(* Logix 5000 project; controller R400_500_XLS vendor 1 type 14 code 216 rev 31.11; software revision 31.01; part 9 of 32 *)
(* tags used below, declared in another part *)
   Abort1 : DINT;   // Not Used
   Alarm : SINT;   // Wait 3 seconds
   Ashutdown : SINT;   // Not Used
   Condenser : INT;
   CondenserHighFlow_1 : BOOL;   // Enables the condenser high flow valve
   CondenserHighFlow_2 : BOOL;   // Enables the condenser high flow valve
   CondenserLowFlow_1 : BOOL;   // Enables the condenser low flow valve
   CondenserLowFlow_2 : BOOL;   // Enables the condenser low flow valve
   CURRENT_CYCLE : DINT;
   CycExcBuffer : UDT_CYCLE;
   Cycles : UDT_CYCLE[11];
   DESCALER : SINT;
   DrnSmp : DINT;
   DRYING : DINT;   // Drying id number
   ENVIRO_CARE : SINT;
   EXTRA_CARE : SINT;
   F1rinse : DINT;   // Not Used
   F2rinse : DINT;   // Not Used
   F3rinse : DINT;   // Not Used
   F4rinse : INT;   // Transition for the conductivity based evalutaion
   FC22_WashIndex : SINT;
   FC23_WashIndex : DINT;   // Current index of the wash treatment
   FC87_CalibChemPmp : SINT;   // Calibration chemical pumps activation bits
   Fill_Sump : DINT;
   HeatSmp : DINT;
   Inj_Cond : SINT;   // Conductivity injection based steps
   Inj_Time : SINT;   // Time based chemical injection steps
   M : DINT[5];   // Memory Bits
   NeutralizantPump : SINT;
   PLASTIC_CARE : SINT;
   PrimeChemPmp : SINT;   // Prime chemical pumps activation bits
   PureWaterTankFilling : BOOL;   // Start PWT filling
   PWR_UP : DINT;
   RINSE_CARE : SINT;
   Run : DINT;
   Service : DINT[2];   // Unused Service Mode Memory Bit
   Shutdown : SINT;   // Shutdown sequence steps
   STANDARD : SINT;
   StartPump1 : BOOL;   // Pump Low Speed
   StartPump2 : BOOL;   // Pump High Speed
   Tmr : TIMER[107];
   Trt_Vapor_Exhaust : BOOL;   // Vapor exhaust fan is on
   USER_DEFINED_10 : SINT;
   USER_DEFINED_11 : SINT;
   USER_DEFINED_7 : SINT;
   USER_DEFINED_8 : SINT;
   USER_DEFINED_9 : SINT;
   AlarmTrigger : INT;   // Triggers the alarm screen if different of 0
   CR2Mode : SINT;   // 0= Cycle complete dry contact 1= External pure water valve
   CycleName : STRING[12];
   CyclePtr : DINT;   // Cycle Pointeur
   I_Pw_Tnk_Sft_Lvl_Sw : BOOL;   // Pure water tank safety level switch
   I_Smp_Sft_Lvl_Sw : BOOL;   // Sump safety level switch
   PureWaterTankDrainingDeadLeg : BOOL;
   Q_Adble_Alrm : BOOL;   // Audible Alarm and /Pilot Light: red connection
   Q_Chm_1 : BOOL;   // Chemical pump #1
   Q_Chm_2 : BOOL;   // Chemical pump #2
   Q_Chm_3 : BOOL;   // Chemical pump #3
   Q_Chm_4 : BOOL;   // Chemical pump #4
   Q_Cld_Wtr_Fll_Vlve : BOOL;   // Cold water sump fill valve
   Q_Cmmn_Alrm : BOOL;   // Dry contact For Alarm
   Q_Cndsr_Hflw_Vlve : BOOL;   // Condenser high flow cold water valve
   Q_Cndsr_Lflw_Vlve : BOOL;   // Condenser low flow cold water valve
   Q_Cyc_Comp : BOOL;   // Dry Contact For Cycle Completed or Pure Water fill valve
   Q_Cyc_Run : BOOL;   // Pilot light: Green connection
   Q_Drn_Cldwn_Vlve : BOOL;   // Drain cool down water valve
   Q_Dry_Fan : BOOL;   // Vapor removal fan / Drying fan
   Q_Dry_Htr : BOOL;   // Drying heating elements
   Q_Dry_Iso_Vlve : BOOL;   // Drying Isolation Valve (Normally Closed Valve)
   Q_Ht_Rcvry_Tnk_Drn_Vlve : BOOL;   // Heat recovery tank drian valve
   Q_Ht_Wtr_Fll_Vlve : BOOL;   // Hot water sump fill valve
   Q_Int_Lght : BOOL;   // Interior Light
   Q_Pmp_Hgh_Spd : BOOL;   // Pump high speed
   Q_Pmp_Lw_Spd : BOOL;   // Pump low speed
   Q_Pw_Fll_Vlve : BOOL;   // Pure water sump/ Tank fill valve
   Q_Pw_Otlt_Vlve : BOOL;   // Pure water tank outlet valve
   Q_Pw_Tnk_Stm_Vlve : BOOL;   // PWT Steam Valve / Electric Heater
   Q_Smp_drn_Vlve : BOOL;   // Sump drain valve (Normally open valve)
   Q_Smp_Stm_Vlve : BOOL;   // Sump steam valve/ Electrical Heater
   Q_Trsfr_Vlve : BOOL;   // Transfer Valve (Normally Open Valve)
   Screen_Ctrl : DINT;   // PLC Screen Request
   Tpb : DINT[11];
   Unit : Hrdwre;   // Unit Configuration
(* MainProgram, continued *)

ROUTINE OPR_9_SELECT_CYCLE   (* ladder *)
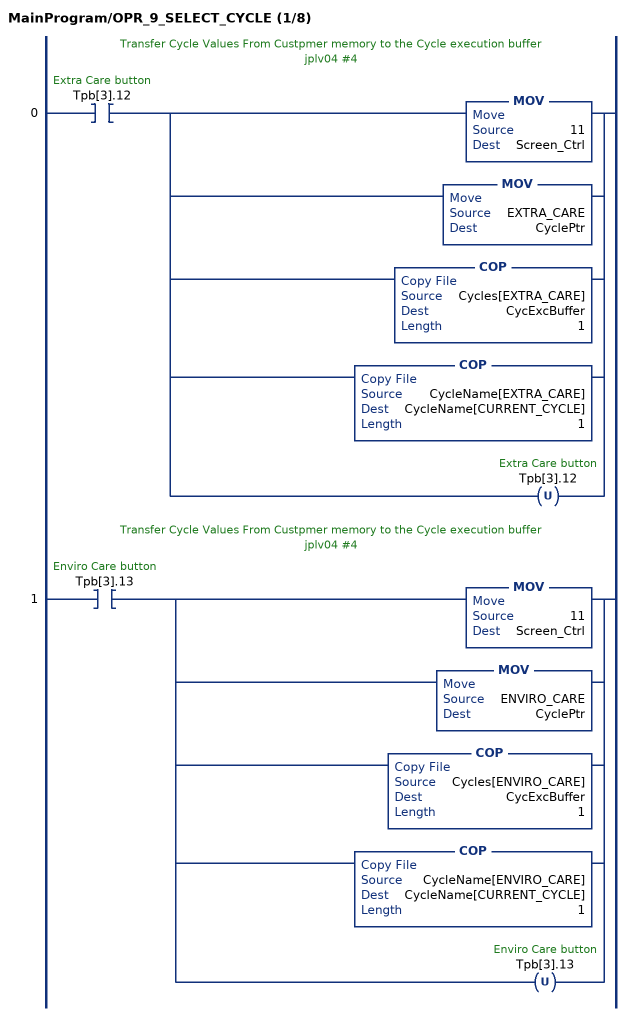
   // Transfer Cycle Values From Custpmer memory to the Cycle execution buffer
   //  jplv04 #4
   0: XIC(Tpb[3].12)[MOV(11,Screen_Ctrl) ,MOV(EXTRA_CARE,CyclePtr) ,COP(Cycles[EXTRA_CARE],CycExcBuffer,1) ,COP(CycleName[EXTRA_CARE],CycleName[CURRENT_CYCLE],1) ,OTU(Tpb[3].12) ];
   // Transfer Cycle Values From Custpmer memory to the Cycle execution buffer
   // jplv04 #4
   1: XIC(Tpb[3].13)[MOV(11,Screen_Ctrl) ,MOV(ENVIRO_CARE,CyclePtr) ,COP(Cycles[ENVIRO_CARE],CycExcBuffer,1) ,COP(CycleName[ENVIRO_CARE],CycleName[CURRENT_CYCLE],1) ,OTU(Tpb[3].13) ];
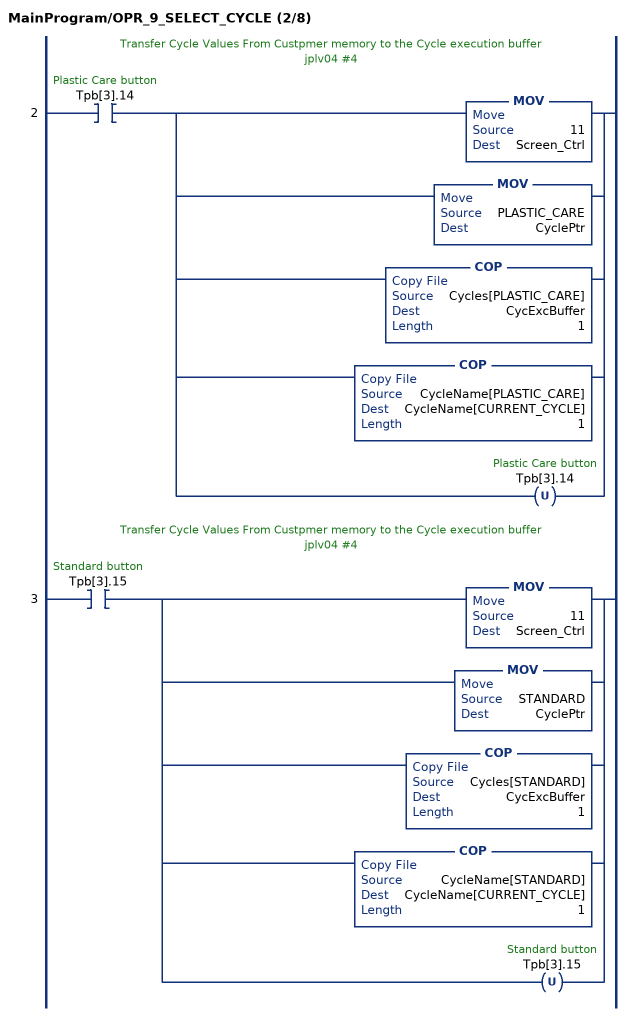
   // Transfer Cycle Values From Custpmer memory to the Cycle execution buffer
   // jplv04 #4
   2: XIC(Tpb[3].14)[MOV(11,Screen_Ctrl) ,MOV(PLASTIC_CARE,CyclePtr) ,COP(Cycles[PLASTIC_CARE],CycExcBuffer,1) ,COP(CycleName[PLASTIC_CARE],CycleName[CURRENT_CYCLE],1) ,OTU(Tpb[3].14) ];
   // Transfer Cycle Values From Custpmer memory to the Cycle execution buffer
   // jplv04 #4
   3: XIC(Tpb[3].15)[MOV(11,Screen_Ctrl) ,MOV(STANDARD,CyclePtr) ,COP(Cycles[STANDARD],CycExcBuffer,1) ,COP(CycleName[STANDARD],CycleName[CURRENT_CYCLE],1) ,OTU(Tpb[3].15) ];
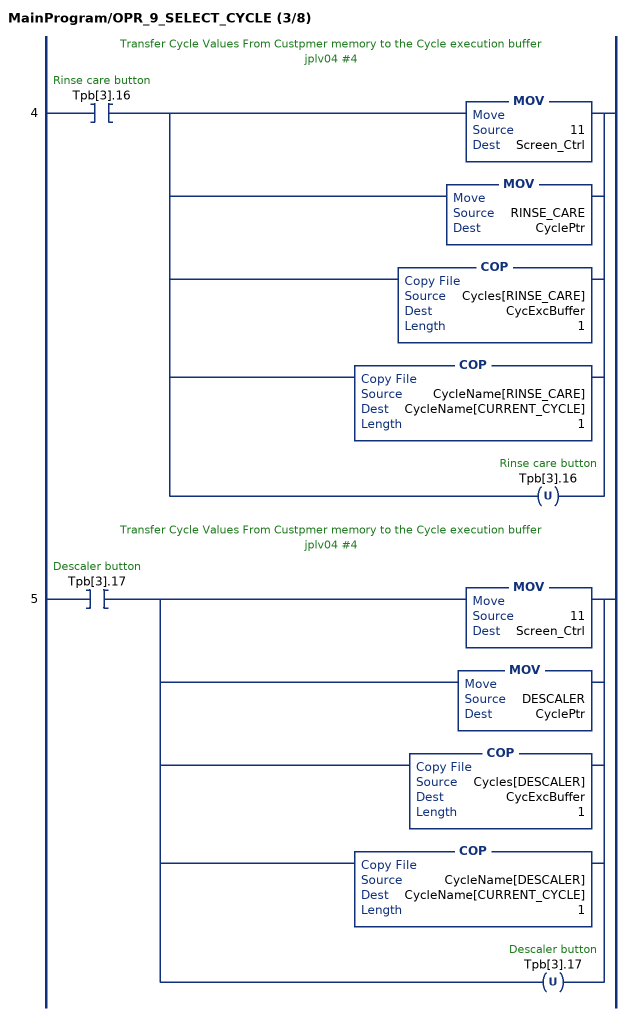
   // Transfer Cycle Values From Custpmer memory to the Cycle execution buffer
   // jplv04 #4
   4: XIC(Tpb[3].16)[MOV(11,Screen_Ctrl) ,MOV(RINSE_CARE,CyclePtr) ,COP(Cycles[RINSE_CARE],CycExcBuffer,1) ,COP(CycleName[RINSE_CARE],CycleName[CURRENT_CYCLE],1) ,OTU(Tpb[3].16) ];
   // Transfer Cycle Values From Custpmer memory to the Cycle execution buffer
   // jplv04 #4
   5: XIC(Tpb[3].17)[MOV(11,Screen_Ctrl) ,MOV(DESCALER,CyclePtr) ,COP(Cycles[DESCALER],CycExcBuffer,1) ,COP(CycleName[DESCALER],CycleName[CURRENT_CYCLE],1) ,OTU(Tpb[3].17) ];
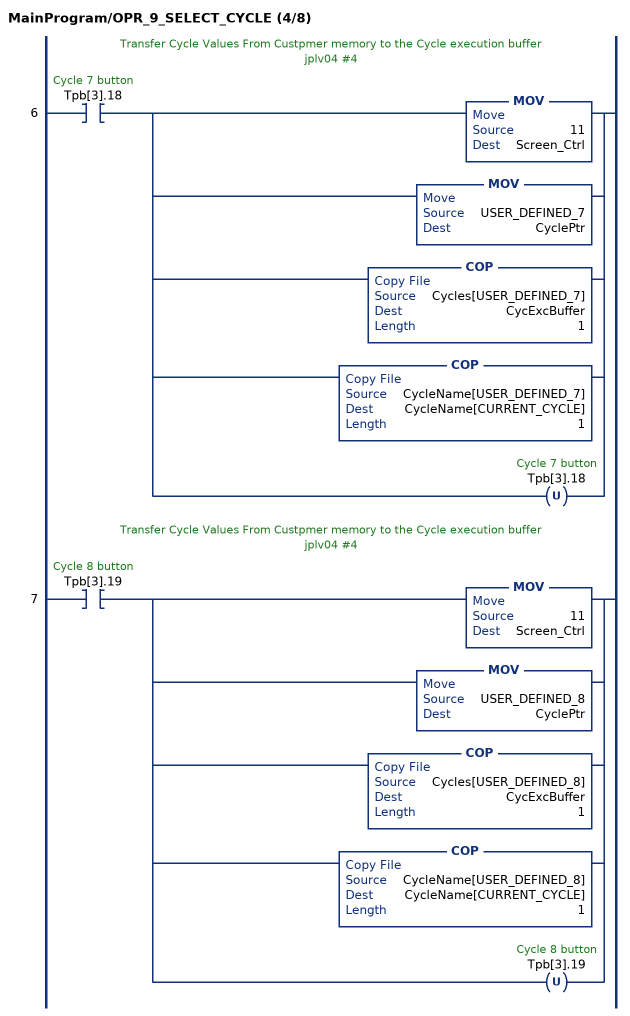
   // Transfer Cycle Values From Custpmer memory to the Cycle execution buffer
   // jplv04 #4
   6: XIC(Tpb[3].18)[MOV(11,Screen_Ctrl) ,MOV(USER_DEFINED_7,CyclePtr) ,COP(Cycles[USER_DEFINED_7],CycExcBuffer,1) ,COP(CycleName[USER_DEFINED_7],CycleName[CURRENT_CYCLE],1) ,OTU(Tpb[3].18) ];
   // Transfer Cycle Values From Custpmer memory to the Cycle execution buffer
   // jplv04 #4
   7: XIC(Tpb[3].19)[MOV(11,Screen_Ctrl) ,MOV(USER_DEFINED_8,CyclePtr) ,COP(Cycles[USER_DEFINED_8],CycExcBuffer,1) ,COP(CycleName[USER_DEFINED_8],CycleName[CURRENT_CYCLE],1) ,OTU(Tpb[3].19) ];
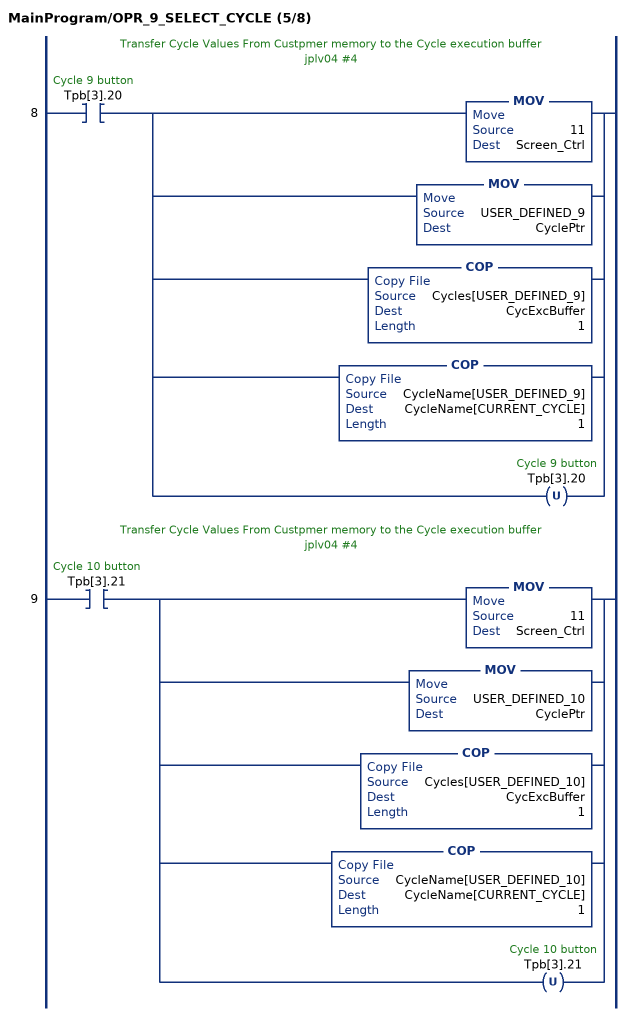
   // Transfer Cycle Values From Custpmer memory to the Cycle execution buffer
   // jplv04 #4
   8: XIC(Tpb[3].20)[MOV(11,Screen_Ctrl) ,MOV(USER_DEFINED_9,CyclePtr) ,COP(Cycles[USER_DEFINED_9],CycExcBuffer,1) ,COP(CycleName[USER_DEFINED_9],CycleName[CURRENT_CYCLE],1) ,OTU(Tpb[3].20) ];
   // Transfer Cycle Values From Custpmer memory to the Cycle execution buffer
   // jplv04 #4
   9: XIC(Tpb[3].21)[MOV(11,Screen_Ctrl) ,MOV(USER_DEFINED_10,CyclePtr) ,COP(Cycles[USER_DEFINED_10],CycExcBuffer,1) ,COP(CycleName[USER_DEFINED_10],CycleName[CURRENT_CYCLE],1) ,OTU(Tpb[3].21) ];
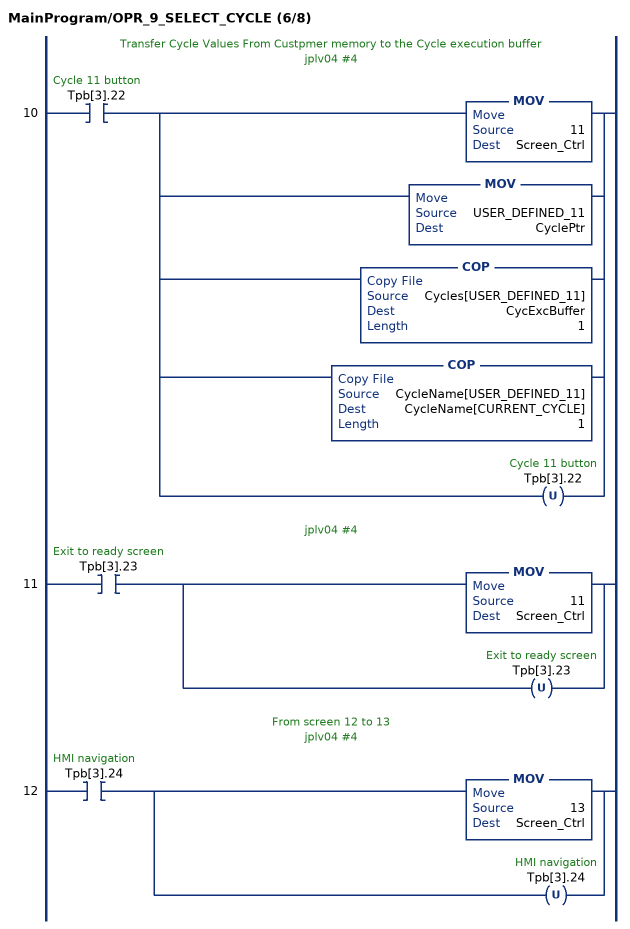
   // Transfer Cycle Values From Custpmer memory to the Cycle execution buffer
   // jplv04 #4
   10: XIC(Tpb[3].22)[MOV(11,Screen_Ctrl) ,MOV(USER_DEFINED_11,CyclePtr) ,COP(Cycles[USER_DEFINED_11],CycExcBuffer,1) ,COP(CycleName[USER_DEFINED_11],CycleName[CURRENT_CYCLE],1) ,OTU(Tpb[3].22) ];
   // jplv04 #4
   11: XIC(Tpb[3].23)[MOV(11,Screen_Ctrl) ,OTU(Tpb[3].23) ];
   // From screen 12 to 13
   // jplv04 #4
   12: XIC(Tpb[3].24)[MOV(13,Screen_Ctrl) ,OTU(Tpb[3].24) ];
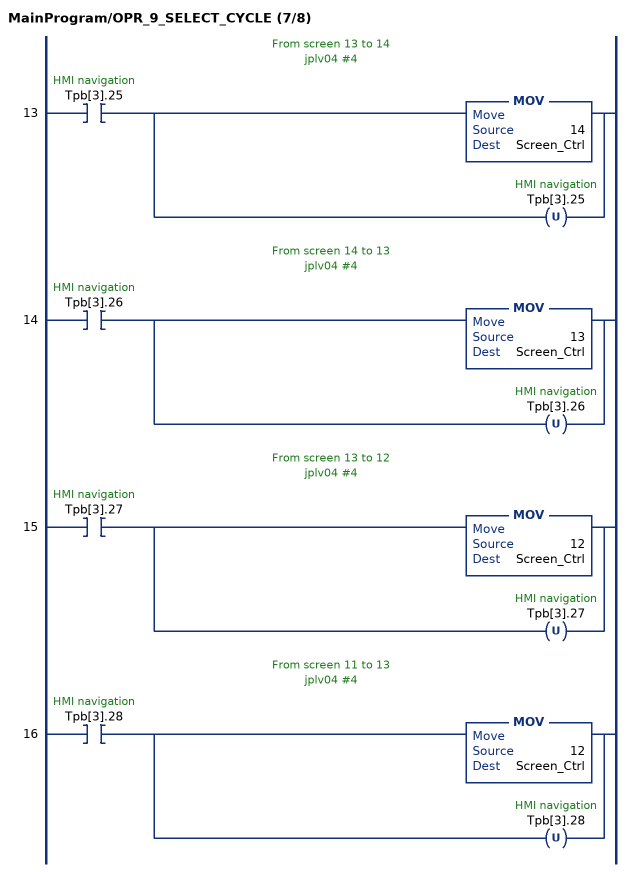
   // From screen 13 to 14
   // jplv04 #4
   13: XIC(Tpb[3].25)[MOV(14,Screen_Ctrl) ,OTU(Tpb[3].25) ];
   // From screen 14 to 13
   // jplv04 #4
   14: XIC(Tpb[3].26)[MOV(13,Screen_Ctrl) ,OTU(Tpb[3].26) ];
   // From screen 13 to 12
   // jplv04 #4
   15: XIC(Tpb[3].27)[MOV(12,Screen_Ctrl) ,OTU(Tpb[3].27) ];
   // From screen 11 to 13
   // jplv04 #4
   16: XIC(Tpb[3].28)[MOV(12,Screen_Ctrl) ,OTU(Tpb[3].28) ];
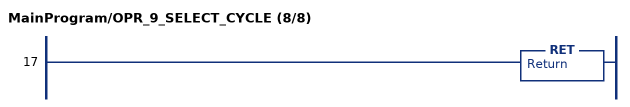
   17: RET();
END_ROUTINE

ROUTINE Outputs   (* ladder *)
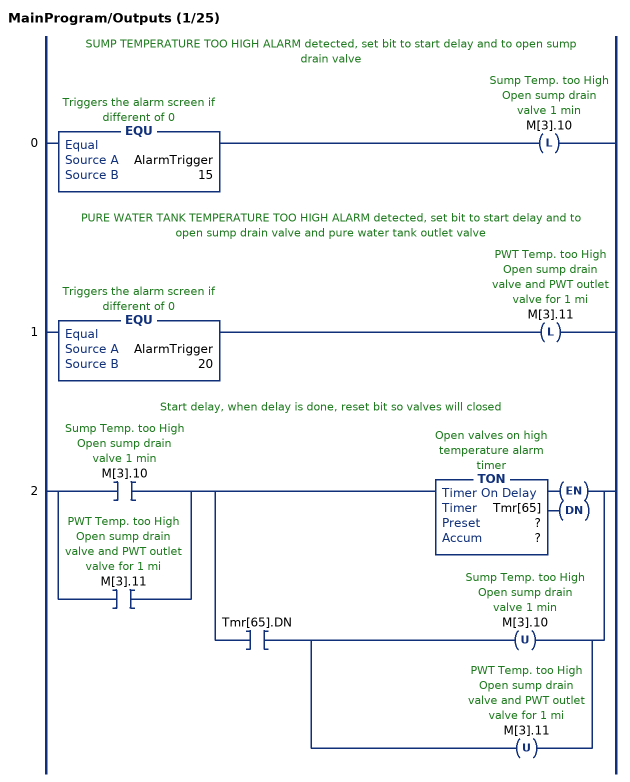
   // SUMP TEMPERATURE TOO HIGH ALARM detected, set bit to start delay and to open sump drain valve
   0: EQU(AlarmTrigger,15)OTL(M[3].10);
   // PURE WATER TANK TEMPERATURE TOO HIGH ALARM detected, set bit to start delay and to open sump drain valve and pure water tank outlet valve
   1: EQU(AlarmTrigger,20)OTL(M[3].11);
   // Start delay, when delay is done, reset bit so valves will closed
   2: [XIC(M[3].10) ,XIC(M[3].11) ][TON(Tmr[65],?,?) ,XIC(Tmr[65].DN) [OTU(M[3].10) ,OTU(M[3].11) ] ];
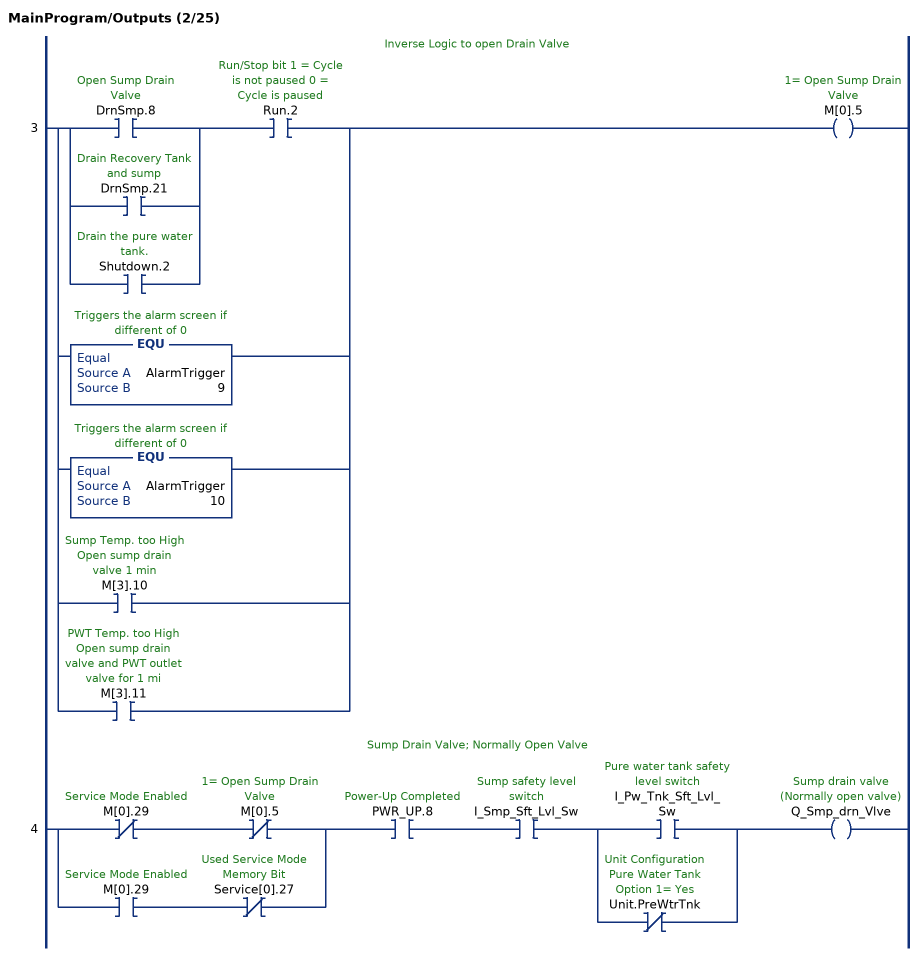
   // Inverse Logic to open Drain Valve
   3: [[XIC(DrnSmp.8) ,XIC(DrnSmp.21) ,XIC(Shutdown.2) ] XIC(Run.2) ,EQU(AlarmTrigger,9) ,EQU(AlarmTrigger,10) ,XIC(M[3].10) ,XIC(M[3].11) ]OTE(M[0].5);
   // Sump Drain Valve; Normally Open Valve
   4: [XIO(M[0].29) XIO(M[0].5) ,XIC(M[0].29) XIO(Service[0].27) ]XIC(PWR_UP.8)XIC(I_Smp_Sft_Lvl_Sw)[XIC(I_Pw_Tnk_Sft_Lvl_Sw) ,XIO(Unit.PreWtrTnk) ]OTE(Q_Smp_drn_Vlve);
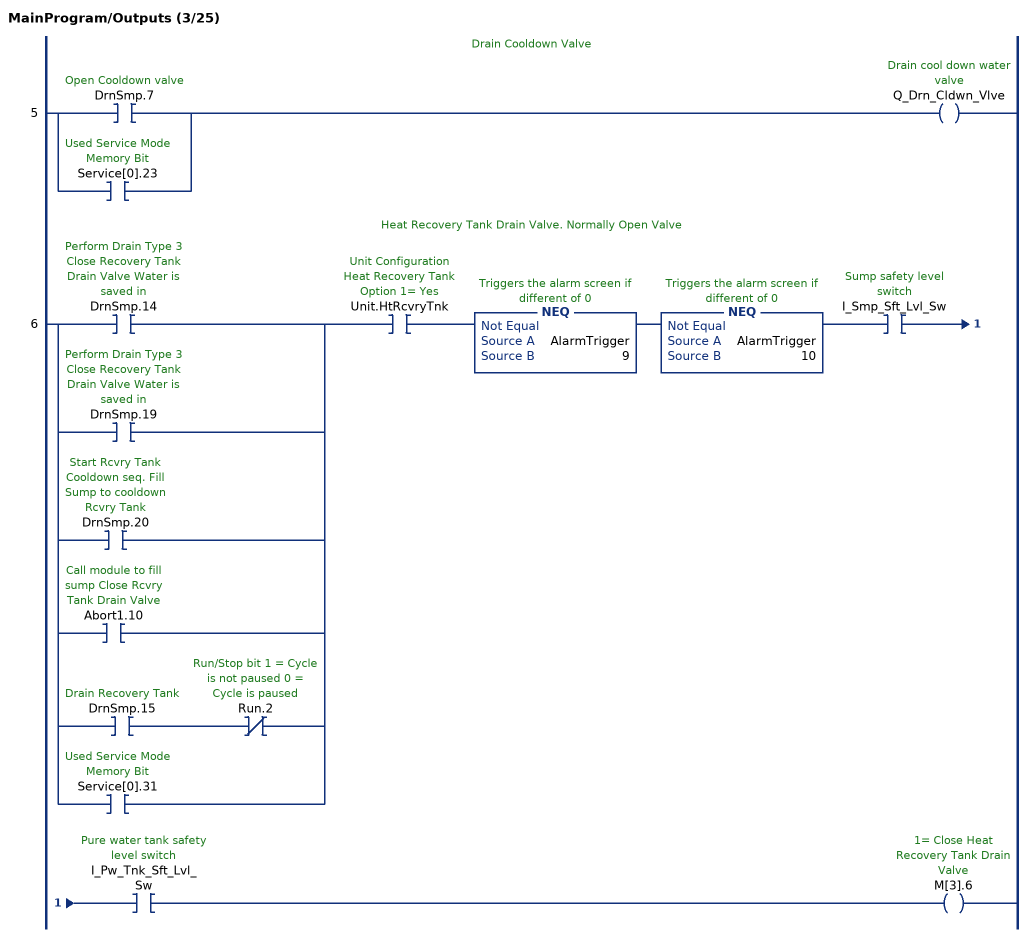
   // Drain Cooldown Valve
   5: [XIC(DrnSmp.7) ,XIC(Service[0].23) ]OTE(Q_Drn_Cldwn_Vlve);
   // Heat Recovery Tank Drain Valve. Normally Open Valve
   6: [XIC(DrnSmp.14) ,XIC(DrnSmp.19) ,XIC(DrnSmp.20) ,XIC(Abort1.10) ,XIC(DrnSmp.15) XIO(Run.2) ,XIC(Service[0].31) ]XIC(Unit.HtRcvryTnk)NEQ(AlarmTrigger,9)NEQ(AlarmTrigger,10)XIC(I_Smp_Sft_Lvl_Sw)XIC(I_Pw_Tnk_Sft_Lvl_Sw)OTE(M[3].6);
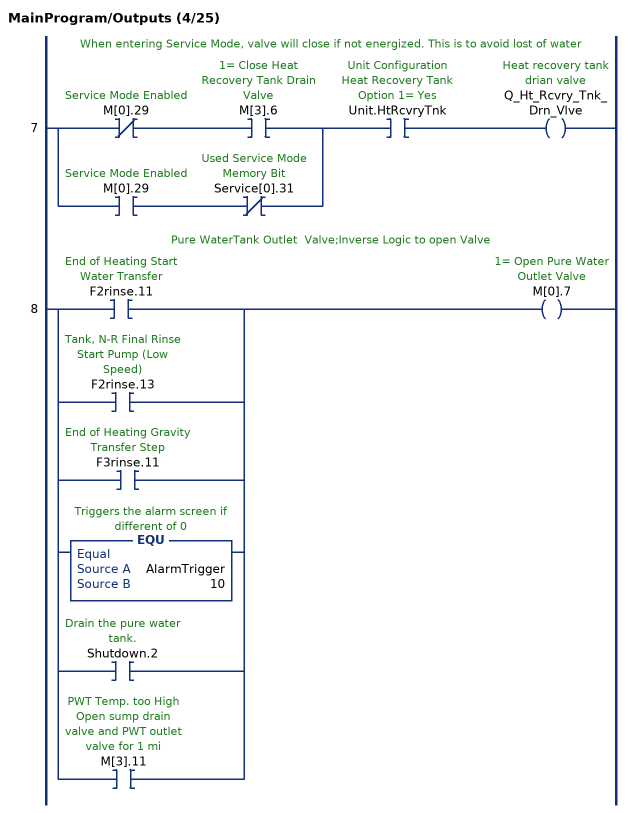
   // When entering Service Mode, valve will close if not energized. This is to avoid lost of water
   7: [XIO(M[0].29) XIC(M[3].6) ,XIC(M[0].29) XIO(Service[0].31) ]XIC(Unit.HtRcvryTnk)OTE(Q_Ht_Rcvry_Tnk_Drn_Vlve);
   // Pure WaterTank Outlet  Valve;Inverse Logic to open Valve
   8: [XIC(F2rinse.11) ,XIC(F2rinse.13) ,XIC(F3rinse.11) ,EQU(AlarmTrigger,10) ,XIC(Shutdown.2) ,XIC(M[3].11) ]OTE(M[0].7);
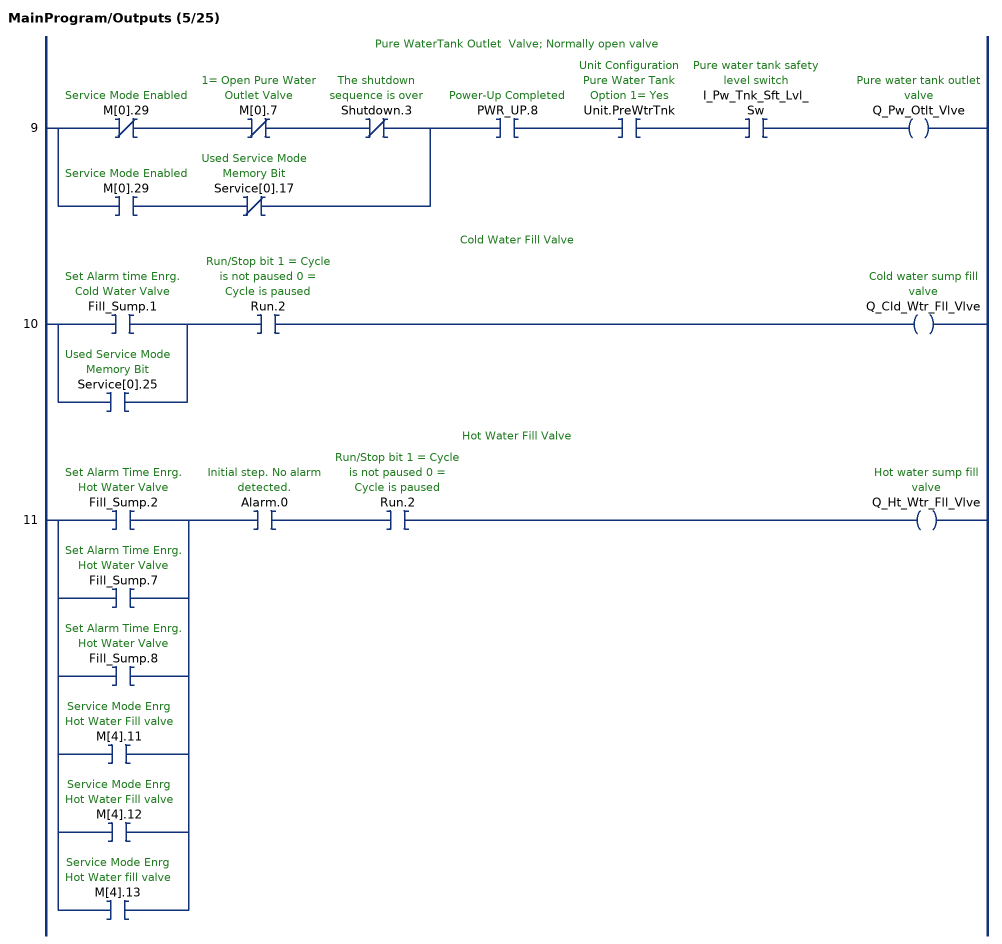
   // Pure WaterTank Outlet  Valve; Normally open valve
   9: [XIO(M[0].29) XIO(M[0].7) XIO(Shutdown.3) ,XIC(M[0].29) XIO(Service[0].17) ]XIC(PWR_UP.8)XIC(Unit.PreWtrTnk)XIC(I_Pw_Tnk_Sft_Lvl_Sw)OTE(Q_Pw_Otlt_Vlve);
   // Cold Water Fill Valve
   10: [XIC(Fill_Sump.1) ,XIC(Service[0].25) ]XIC(Run.2)OTE(Q_Cld_Wtr_Fll_Vlve);
   // Hot Water Fill Valve
   11: [XIC(Fill_Sump.2) ,XIC(Fill_Sump.7) ,XIC(Fill_Sump.8) ,XIC(M[4].11) ,XIC(M[4].12) ,XIC(M[4].13) ]XIC(Alarm.0)XIC(Run.2)OTE(Q_Ht_Wtr_Fll_Vlve);
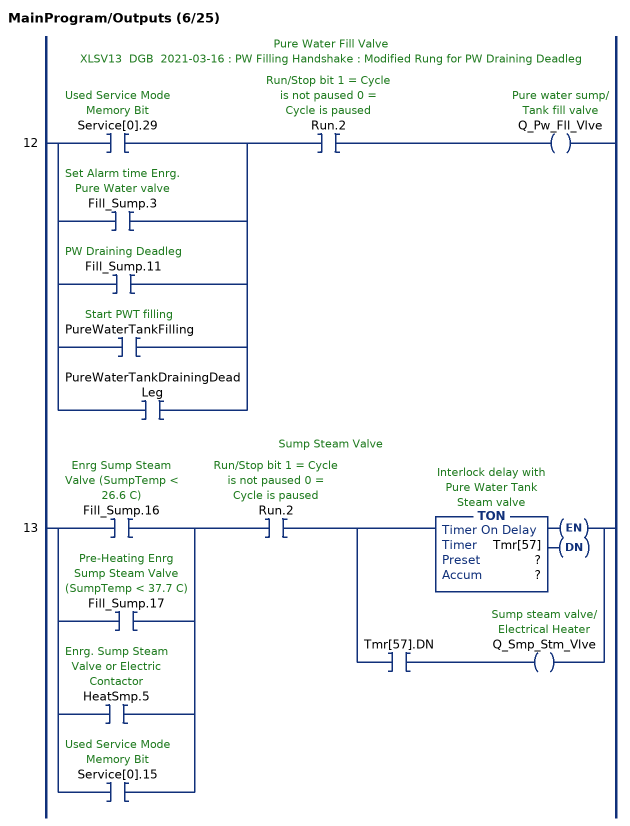
   // Pure Water Fill Valve
   // XLSV13  DGB  2021-03-16 : PW Filling Handshake : Modified Rung for PW Draining Deadleg
   12: [XIC(Service[0].29) ,XIC(Fill_Sump.3) ,XIC(Fill_Sump.11) ,XIC(PureWaterTankFilling) ,XIC(PureWaterTankDrainingDeadLeg) ]XIC(Run.2)OTE(Q_Pw_Fll_Vlve);
   // Sump Steam Valve
   13: [XIC(Fill_Sump.16) ,XIC(Fill_Sump.17) ,XIC(HeatSmp.5) ,XIC(Service[0].15) ]XIC(Run.2)[TON(Tmr[57],?,?) ,XIC(Tmr[57].DN) OTE(Q_Smp_Stm_Vlve) ];
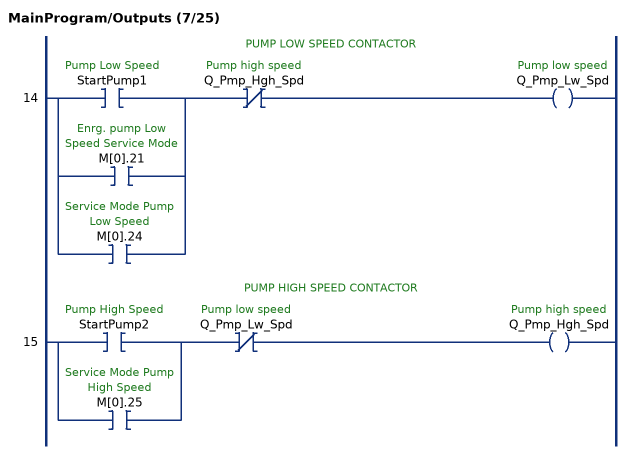
   // PUMP LOW SPEED CONTACTOR
   14: [XIC(StartPump1) ,XIC(M[0].21) ,XIC(M[0].24) ]XIO(Q_Pmp_Hgh_Spd)OTE(Q_Pmp_Lw_Spd);
   // PUMP HIGH SPEED CONTACTOR
   15: [XIC(StartPump2) ,XIC(M[0].25) ]XIO(Q_Pmp_Lw_Spd)OTE(Q_Pmp_Hgh_Spd);
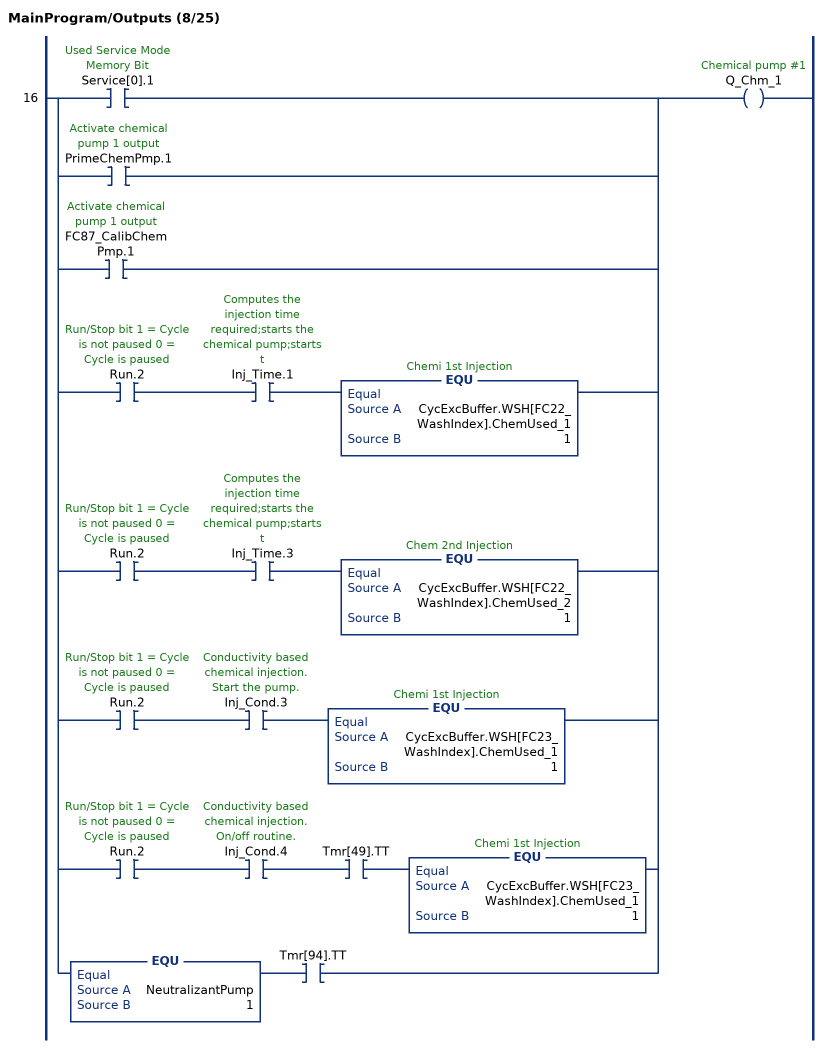
   16: [XIC(Service[0].1) ,XIC(PrimeChemPmp.1) ,XIC(FC87_CalibChemPmp.1) ,XIC(Run.2) XIC(Inj_Time.1) EQU(CycExcBuffer.WSH[FC22_WashIndex].ChemUsed_1,1) ,XIC(Run.2) XIC(Inj_Time.3) EQU(CycExcBuffer.WSH[FC22_WashIndex].ChemUsed_2,1) ,XIC(Run.2) XIC(Inj_Cond.3) EQU(CycExcBuffer.WSH[FC23_WashIndex].ChemUsed_1,1) ,XIC(Run.2) XIC(Inj_Cond.4) XIC(Tmr[49].TT) EQU(CycExcBuffer.WSH[FC23_WashIndex].ChemUsed_1,1) ,EQU(NeutralizantPump,1) XIC(Tmr[94].TT) ]OTE(Q_Chm_1);
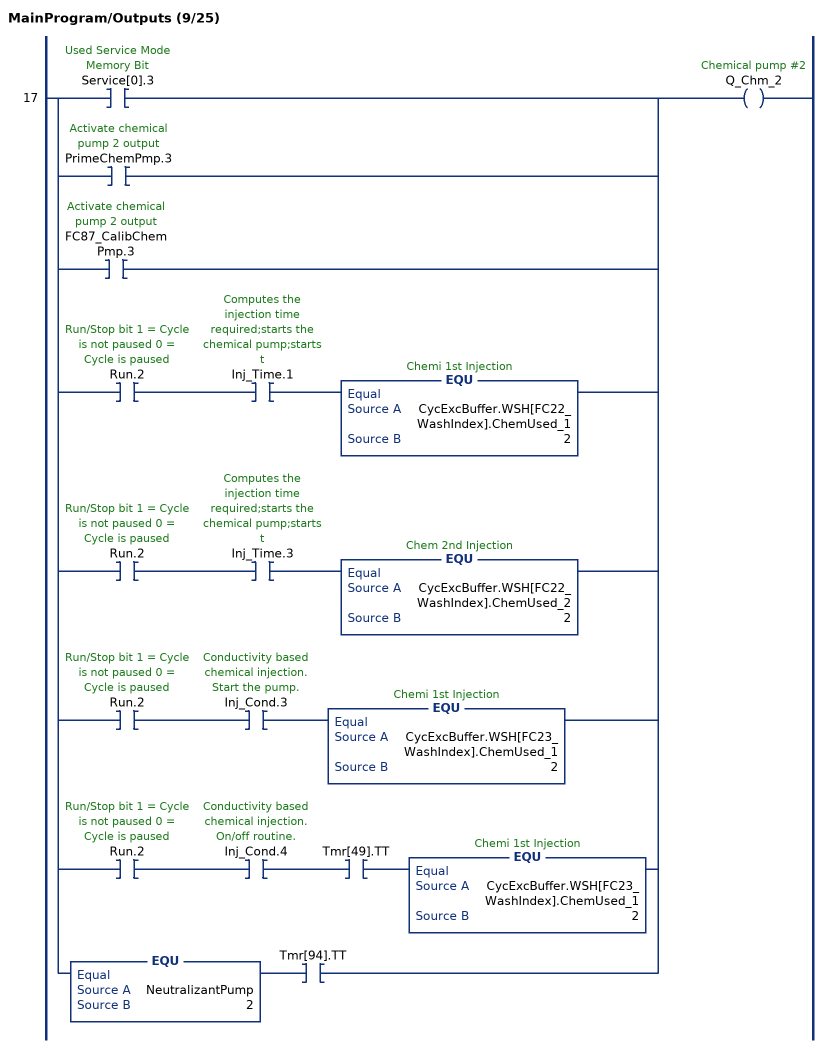
   17: [XIC(Service[0].3) ,XIC(PrimeChemPmp.3) ,XIC(FC87_CalibChemPmp.3) ,XIC(Run.2) XIC(Inj_Time.1) EQU(CycExcBuffer.WSH[FC22_WashIndex].ChemUsed_1,2) ,XIC(Run.2) XIC(Inj_Time.3) EQU(CycExcBuffer.WSH[FC22_WashIndex].ChemUsed_2,2) ,XIC(Run.2) XIC(Inj_Cond.3) EQU(CycExcBuffer.WSH[FC23_WashIndex].ChemUsed_1,2) ,XIC(Run.2) XIC(Inj_Cond.4) XIC(Tmr[49].TT) EQU(CycExcBuffer.WSH[FC23_WashIndex].ChemUsed_1,2) ,EQU(NeutralizantPump,2) XIC(Tmr[94].TT) ]OTE(Q_Chm_2);
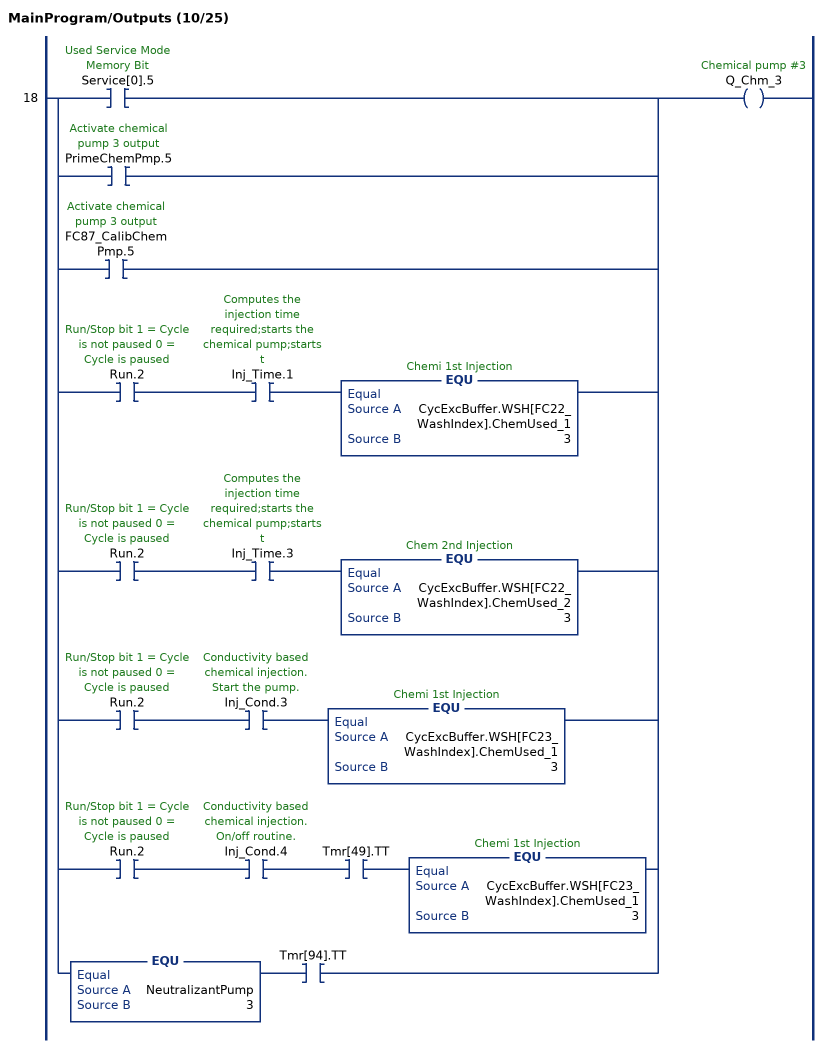
   18: [XIC(Service[0].5) ,XIC(PrimeChemPmp.5) ,XIC(FC87_CalibChemPmp.5) ,XIC(Run.2) XIC(Inj_Time.1) EQU(CycExcBuffer.WSH[FC22_WashIndex].ChemUsed_1,3) ,XIC(Run.2) XIC(Inj_Time.3) EQU(CycExcBuffer.WSH[FC22_WashIndex].ChemUsed_2,3) ,XIC(Run.2) XIC(Inj_Cond.3) EQU(CycExcBuffer.WSH[FC23_WashIndex].ChemUsed_1,3) ,XIC(Run.2) XIC(Inj_Cond.4) XIC(Tmr[49].TT) EQU(CycExcBuffer.WSH[FC23_WashIndex].ChemUsed_1,3) ,EQU(NeutralizantPump,3) XIC(Tmr[94].TT) ]OTE(Q_Chm_3);
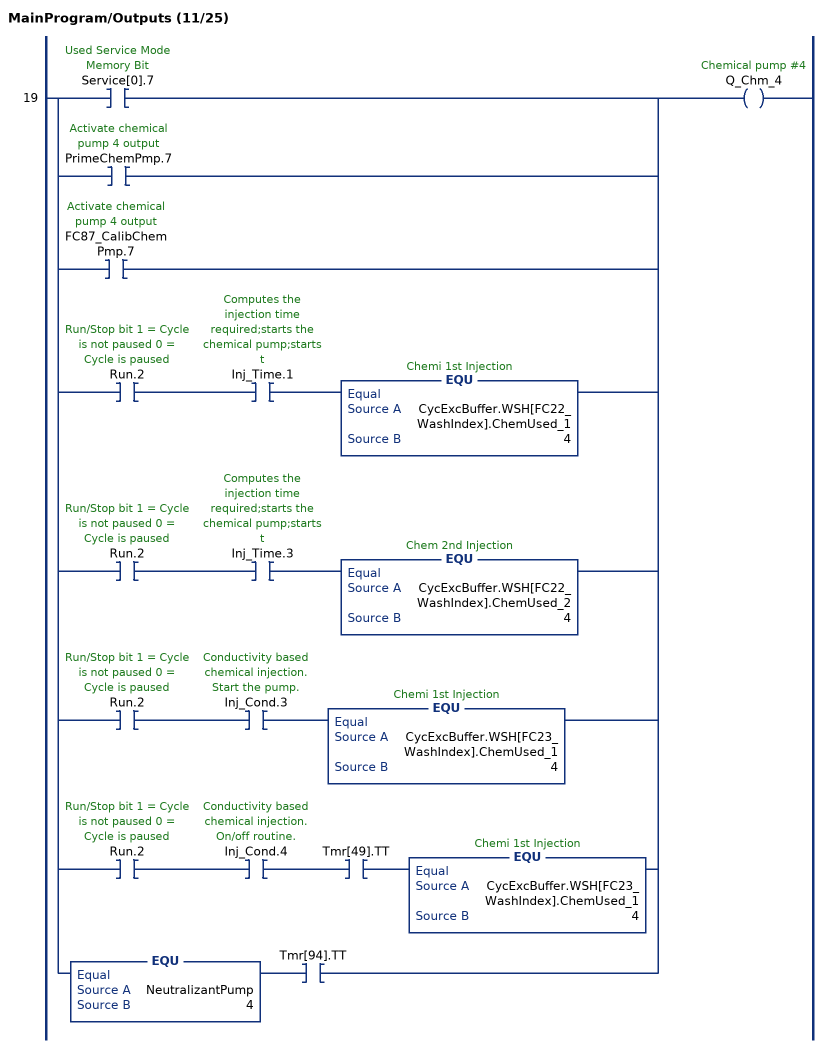
   19: [XIC(Service[0].7) ,XIC(PrimeChemPmp.7) ,XIC(FC87_CalibChemPmp.7) ,XIC(Run.2) XIC(Inj_Time.1) EQU(CycExcBuffer.WSH[FC22_WashIndex].ChemUsed_1,4) ,XIC(Run.2) XIC(Inj_Time.3) EQU(CycExcBuffer.WSH[FC22_WashIndex].ChemUsed_2,4) ,XIC(Run.2) XIC(Inj_Cond.3) EQU(CycExcBuffer.WSH[FC23_WashIndex].ChemUsed_1,4) ,XIC(Run.2) XIC(Inj_Cond.4) XIC(Tmr[49].TT) EQU(CycExcBuffer.WSH[FC23_WashIndex].ChemUsed_1,4) ,EQU(NeutralizantPump,4) XIC(Tmr[94].TT) ]OTE(Q_Chm_4);
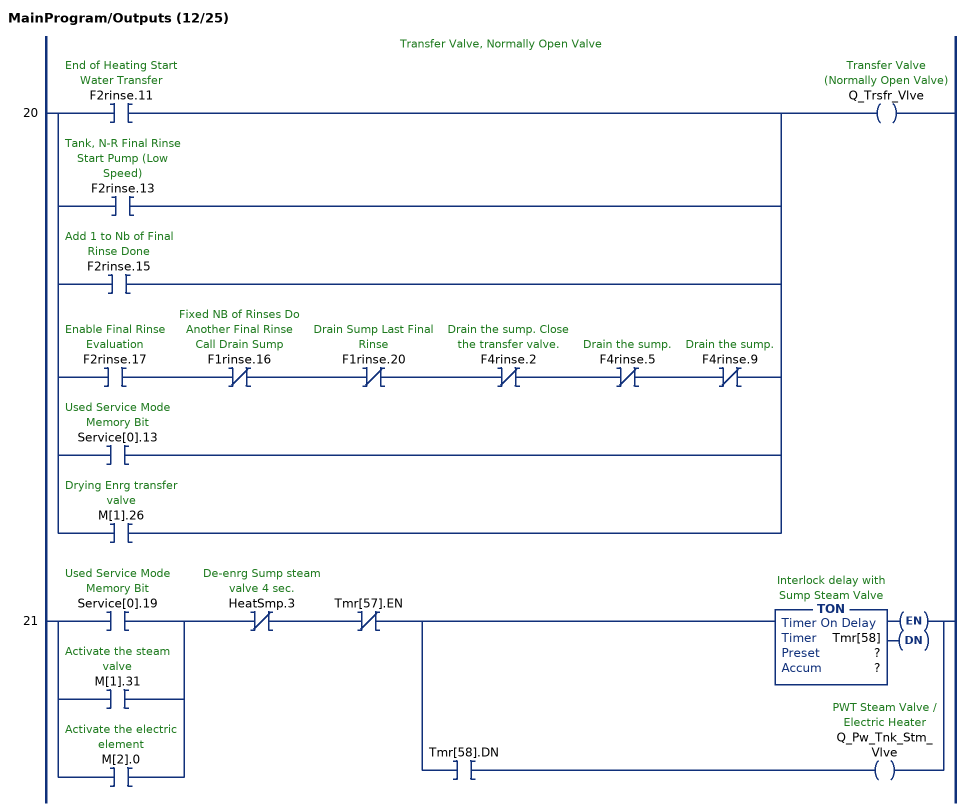
   // Transfer Valve, Normally Open Valve
   20: [[XIC(F2rinse.11) ,XIC(F2rinse.13) ,XIC(F2rinse.15) ,XIC(F2rinse.17) XIO(F1rinse.16) XIO(F1rinse.20) XIO(F4rinse.2) XIO(F4rinse.5) XIO(F4rinse.9) ] ,XIC(Service[0].13) ,XIC(M[1].26) ]OTE(Q_Trsfr_Vlve);
   21: [XIC(Service[0].19) ,XIC(M[1].31) ,XIC(M[2].0) ]XIO(HeatSmp.3)XIO(Tmr[57].EN)[TON(Tmr[58],?,?) ,XIC(Tmr[58].DN) OTE(Q_Pw_Tnk_Stm_Vlve) ];
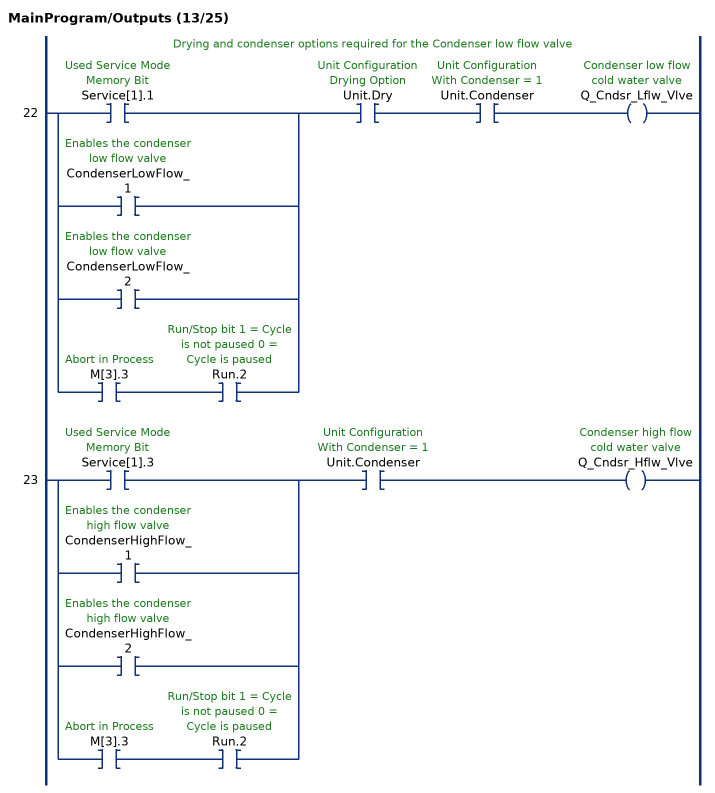
   // Drying and condenser options required for the Condenser low flow valve
   22: [XIC(Service[1].1) ,XIC(CondenserLowFlow_1) ,XIC(CondenserLowFlow_2) ,XIC(M[3].3) XIC(Run.2) ]XIC(Unit.Dry)XIC(Unit.Condenser)OTE(Q_Cndsr_Lflw_Vlve);
   23: [XIC(Service[1].3) ,XIC(CondenserHighFlow_1) ,XIC(CondenserHighFlow_2) ,XIC(M[3].3) XIC(Run.2) ]XIC(Unit.Condenser)OTE(Q_Cndsr_Hflw_Vlve);
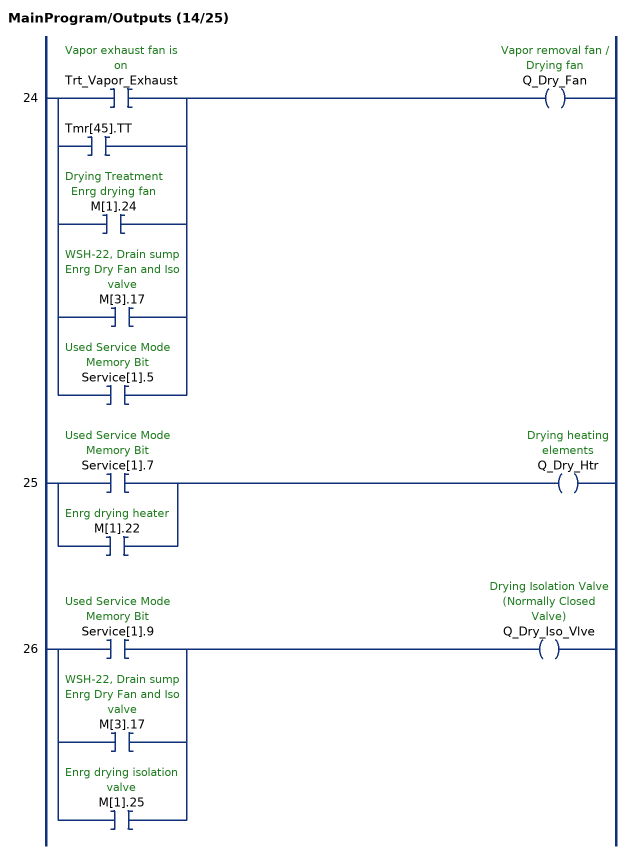
   24: [XIC(Trt_Vapor_Exhaust) ,XIC(Tmr[45].TT) ,XIC(M[1].24) ,XIC(M[3].17) ,XIC(Service[1].5) ]OTE(Q_Dry_Fan);
   25: [XIC(Service[1].7) ,XIC(M[1].22) ]OTE(Q_Dry_Htr);
   26: [XIC(Service[1].9) ,XIC(M[3].17) ,XIC(M[1].25) ]OTE(Q_Dry_Iso_Vlve);
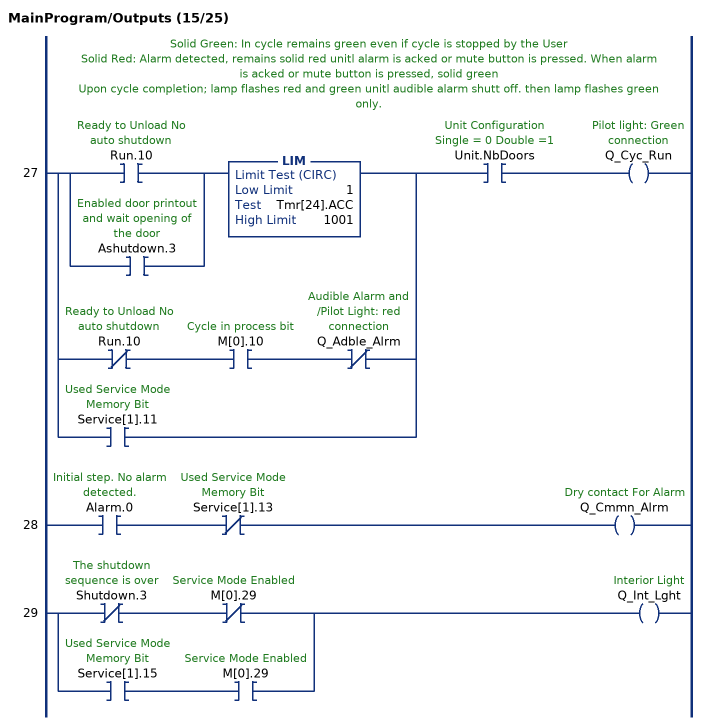
   // Solid Green: In cycle remains green even if cycle is stopped by the User
   // Solid Red: Alarm detected, remains solid red unitl alarm is acked or mute button is pressed. When alarm is acked or mute button is pressed, solid green
   // Upon cycle completion; lamp flashes red and green unitl audible alarm shutt off. then lamp flashes green only.
   27: [[[XIC(Run.10) ,XIC(Ashutdown.3) ] LIM(1,Tmr[24].ACC,1001) ,XIO(Run.10) XIC(M[0].10) XIO(Q_Adble_Alrm) ] ,XIC(Service[1].11) ]XIC(Unit.NbDoors)OTE(Q_Cyc_Run);
   28: XIC(Alarm.0)XIO(Service[1].13)OTE(Q_Cmmn_Alrm);
   29: [XIO(Shutdown.3) XIO(M[0].29) ,XIC(Service[1].15) XIC(M[0].29) ]OTE(Q_Int_Lght);
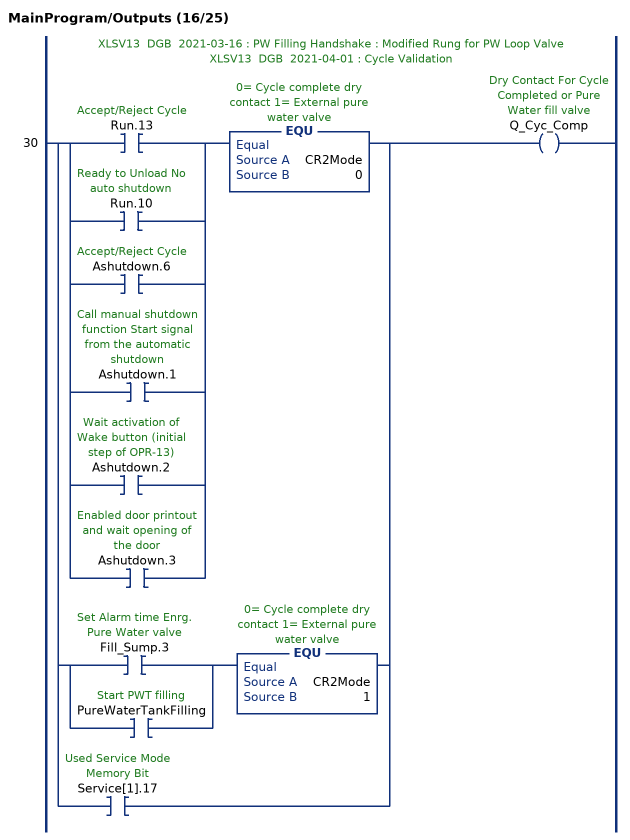
   // XLSV13  DGB  2021-03-16 : PW Filling Handshake : Modified Rung for PW Loop Valve
   // XLSV13  DGB  2021-04-01 : Cycle Validation
   30: [[[XIC(Run.13) ,XIC(Run.10) ,XIC(Ashutdown.6) ,XIC(Ashutdown.1) ,XIC(Ashutdown.2) ,XIC(Ashutdown.3) ] EQU(CR2Mode,0) ,[XIC(Fill_Sump.3) ,XIC(PureWaterTankFilling) ] EQU(CR2Mode,1) ] ,XIC(Service[1].17) ]OTE(Q_Cyc_Comp);
